// TIA Portal V21 export
// export: Created 2026-11-02T00:47:44.0429899Z, ExportSetting WithDefaults, DisplayName Totally Integrated Automation Portal, DisplayVersion V21 Update 3, DisplayName TIA Portal Test Suite Advanced, DisplayVersion V21 Update 1, DisplayName SINAMICS Startdrive Advanced, DisplayVersion V21 Update 1, DisplayName SINAMICS Startdrive G130, G150, S120, S150, G200, G210, G210C, G210X, G220, S200, S210, S220, Innomotics MVD, DisplayVersion V21 Update 1, DisplayName SINAMICS Startdrive G110M, G120, G120C, G120D, G120P, G115D, DisplayVersion V21 Update 1, DisplayName STEP 7 Professional, DisplayVersion V21 Update 3, DisplayName STEP 7 Safety, DisplayVersion V21, DisplayName Tech WebApplication, DisplayVersion V21, DisplayName WinCC Basic/Comfort/Advanced, DisplayVersion V21 Update 3, DisplayName WinCC Professional, DisplayVersion V21 Update 3, DisplayName WinCC Unified, DisplayVersion V21 Update 3
DATA_BLOCK "Tgp_GlobalTemplateFB_LAD"   // DB2
VERSION : 0.1
// stored: AutoNumber true, DBAccessibleFromOPCUA true, DBAccessibleFromWebserver true, InstanceOfName Tgp_TemplateFB_LAD, InstanceOfType FB
"Tgp_TemplateFB_LAD"
   // VAR_INPUT
   //    InputBool : Bool;
   //    InputSInt : SInt;
   //    InputInt : Int;
   //    InputDInt : DInt;
   //    InputLInt : LInt;
   //    InputUSInt : USInt;
   //    InputUInt : UInt;
   //    InputUDInt : UDInt;
   //    InputULInt : ULInt;
   //    InputReal : Real;
   //    InputLReal : LReal;
   //    InputByte : Byte;
   //    InputWord : Word;
   //    InputDWord : DWord;
   //    InputLWord : LWord;
   //    InputTime : Time;
   //    InputLTime : LTime;
   // END_VAR
   // VAR_OUTPUT
   //    OutputBool : Bool;
   //    OutputSInt : SInt;
   //    OutputInt : Int;
   //    OutputDInt : DInt;
   //    OutputLInt : LInt;
   //    OutputUSInt : USInt;
   //    OutputUInt : UInt;
   //    OutputUDInt : UDInt;
   //    OutputULInt : ULInt;
   //    OutputReal : Real;
   //    OutputLReal : LReal;
   //    OutputByte : Byte;
   //    OutputWord : Word;
   //    OutputDWord : DWord;
   //    OutputLWord : LWord;
   //    OutputTime : Time;
   //    OutputLTime : LTime;
   // END_VAR
   // VAR_IN_OUT
   //    InOutBool : Bool;
   //    InOutSInt : SInt;
   //    InOutInt : Int;
   //    InOutDInt : DInt;
   //    InOutLInt : LInt;
   //    InOutUSInt : USInt;
   //    InOutUInt : UInt;
   //    InOutUDInt : UDInt;
   //    InOutULInt : ULInt;
   //    InOutReal : Real;
   //    InOutLReal : LReal;
   //    InOutByte : Byte;
   //    InOutWord : Word;
   //    InOutDWord : DWord;
   //    InOutLWord : LWord;
   //    InOutTime : Time;
   //    InOutLTime : LTime;
   // END_VAR
   // VAR
   //    StaticBool : Bool;
   //    StaticSInt : SInt;
   //    StaticInt : Int;
   //    StaticDInt : DInt;
   //    StaticLInt : LInt;
   //    StaticUSInt : USInt;
   //    StaticUInt : UInt;
   //    StaticUDInt : UDInt;
   //    StaticULInt : ULInt;
   //    StaticReal : Real;
   //    StaticLReal : LReal;
   //    StaticByte : Byte;
   //    StaticWord : Word;
   //    StaticDWord : DWord;
   //    StaticLWord : LWord;
   //    StaticTime : Time;
   //    StaticLTime : LTime;
   // END_VAR
BEGIN
END_DATA_BLOCK
